FUNCTION_BLOCK FB_LintTest EXTENDS FB_LintBase IMPLEMENTS I_LintItf
VAR_INPUT
END_VAR
VAR_OUTPUT
END_VAR
VAR
	nVal : INT;
	sTxt : STRING(40);
END_VAR

nVal := nVal + 1;
A_Act();

ACTION A_Act:
sTxt := 'a]]>b'; // CDATA end marker inside code
END_ACTION

ACTION A_Sfc:
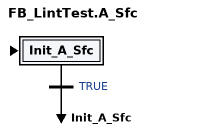
INITIAL_STEP Init_A_Sfc:
END_STEP
TRANSITION FROM Init_A_Sfc TO Init_A_Sfc
    := TRUE;
END_TRANSITION
END_ACTION

METHOD PUBLIC M_Do : BOOL
M_Do := TRUE;
END_METHOD

PROPERTY PUBLIC P_Ro : INT
GET // PUBLIC
P_Ro := 1;
END_GET
END_PROPERTY

PROPERTY PUBLIC P_Val : INT
GET // PUBLIC
P_Val := nVal;
END_GET
SET // PUBLIC
nVal := P_Val;
END_SET
END_PROPERTY

END_FUNCTION_BLOCK

(* stored: Version 1.1.0.1, ProductVersion 3.1.4026.18
   POU FB_LintTest: Id {89e01a82-da3d-04f2-35db-0961eae9f58b}, SpecialFunc None
   Action A_Act: Id {b573562d-f06c-08d5-24b3-b0c2ac52f595}
   Action A_Sfc: Id {f87caa9e-02ca-0868-01e3-07f0d6d66dc6}
   Method M_Do: Id {d9de36ce-09f8-0e34-0bb5-1a4d81e34d82}
   Property P_Ro: Id {50d3f02b-d361-0683-19d1-7d19c7365f0d}
   Get Get: Id {7104f2b8-1acd-0eab-162b-9281c0626913}
   Property P_Val: Id {370cd65e-9ceb-0cd9-33c3-ff0db5ed8e66}
   Get Get: Id {02b0b212-2e05-09dd-0316-862e5c59e067}
   Set Set: Id {a85df9d2-4730-0558-15ff-e6f0c8f709d8} *)
